Fanuc KAREL source: kb00161.KL

-- PROVISIONAL review KL for V1013-1; original PC SHA256 0da0efeac3e0a4bdb45e4160227d7b8c7088bb1fced3043e9094bf0a153fe932
-- Incomplete behavior may be omitted. Consult companion uncertainty JSON. Do not deploy.
PROGRAM KB00161
%NOLOCKGROUP
BEGIN
  -- UNRESOLVED_PC offsets 5-12; opcodes 9D,23
  -- UNRESOLVED_PC offsets 17-24; opcodes 9D,23
  -- UNRESOLVED_PC offsets 29-59; opcodes 27,22,22,1C,22,27,9D,31
  -- UNRESOLVED_PC offsets 64-68; opcodes 7F
END KB00161
